Fanuc KAREL source: KX00015.KL

PROGRAM KX00015
%NOLOCKGROUP
VAR
  I: INTEGER
  J: INTEGER
  B: BOOLEAN
  F: FILE
  S: STRING[80]
  P: XYZWPR
BEGIN
  DISABLE CONDITION[1]
END KX00015
